(* IEC 61131-3 sources: rusty/tests/lit/single/polymorphism/interfaces/properties, 10 files *)

(* ---- basic_get_set.st ---- *)
// RUN: %COMPILE %s && %RUN | %CHECK %s
// Scenario: Single interface with a property declaring both PROPERTY_GET and PROPERTY_SET, implemented by a single
// function block. Assign the concrete instance to an interface variable and exercise both accessors
// through it. Baseline sanity test for property dispatch through interfaces.

INTERFACE IValue
    PROPERTY_GET value: DINT END_PROPERTY
    PROPERTY_SET value: DINT END_PROPERTY
END_INTERFACE

FUNCTION_BLOCK FbStore IMPLEMENTS IValue
    VAR
        _val : DINT := 10;
    END_VAR

    PROPERTY_GET value: DINT
        value := _val;
    END_PROPERTY

    PROPERTY_SET value: DINT
        _val := value;
    END_PROPERTY
END_FUNCTION_BLOCK

FUNCTION main
    VAR
        instance : FbStore;
        iface : IValue;
    END_VAR

    iface := instance;

    // CHECK: value=10
    printf('value=%d$N', iface.value);

    iface.value := 42;

    // CHECK-NEXT: value=42
    printf('value=%d$N', iface.value);

    iface.value := iface.value + 8;

    // CHECK-NEXT: value=50
    printf('value=%d$N', iface.value);
END_FUNCTION

(* ---- deep_chain_alternating_overrides.st ---- *)
// RUN: %COMPILE %s && %RUN | %CHECK %s
// Scenario: Three-level POU chain FbC → FbB → FbA, where FbA implements IValue. FbB overrides
// only the getter (adds 1000), FbC overrides only the setter (adds 2000). Dispatch through the
// interface should resolve each accessor to the most-derived override:
//   FbA → (FbA.get, FbA.set)
//   FbB → (FbB.get, FbA.set)
//   FbC → (FbB.get, FbC.set)

INTERFACE IValue
    PROPERTY_GET value: DINT END_PROPERTY
    PROPERTY_SET value: DINT END_PROPERTY
END_INTERFACE

FUNCTION_BLOCK FbA IMPLEMENTS IValue
    VAR
        _val : DINT := 10;
    END_VAR

    PROPERTY_GET value: DINT
        value := _val;
    END_PROPERTY

    PROPERTY_SET value: DINT
        _val := value;
    END_PROPERTY
END_FUNCTION_BLOCK

FUNCTION_BLOCK FbB EXTENDS FbA
    // Override only getter — adds 1000
    PROPERTY_GET value: DINT
        value := _val + 1000;
    END_PROPERTY
END_FUNCTION_BLOCK

FUNCTION_BLOCK FbC EXTENDS FbB
    // Override only setter — adds 2000
    PROPERTY_SET value: DINT
        _val := value + 2000;
    END_PROPERTY
END_FUNCTION_BLOCK

FUNCTION main
    VAR
        instanceA : FbA;
        instanceB : FbB;
        instanceC : FbC;
        iface : IValue;
    END_VAR

    // FbA: get=FbA, set=FbA
    iface := instanceA;
    printf('value=%d$N', iface.value);      // CHECK: value=10
    iface.value := 50;
    printf('value=%d$N', iface.value);      // CHECK-NEXT: value=50

    // FbB: get=FbB(+1000), set=FbA(inherited)
    iface := instanceB;
    printf('value=%d$N', iface.value);      // CHECK-NEXT: value=1010
    iface.value := 50;
    printf('value=%d$N', iface.value);      // CHECK-NEXT: value=1050

    // FbC: get=FbB(inherited, +1000), set=FbC(+2000)
    iface := instanceC;
    printf('value=%d$N', iface.value);      // CHECK-NEXT: value=1010
    iface.value := 50;
    printf('value=%d$N', iface.value);      // CHECK-NEXT: value=3050
END_FUNCTION

(* ---- diamond_hierarchy.st ---- *)
// RUN: %COMPILE %s && %RUN | %CHECK %s
// Scenario: Classic diamond pattern with a property at the root.
//     IA (property value)
//    /  \
//   IB   IC
//    \  /
//     ID
// IB adds method bar, IC adds method baz, ID adds method qux. A single function block
// FbImpl implements ID (and thus transitively IA, IB, IC). Dispatch through IA, IB, IC
// and ID variables should all resolve the property correctly, and each interface level
// should expose its respective methods.

INTERFACE IA
    PROPERTY_GET value: DINT END_PROPERTY
    PROPERTY_SET value: DINT END_PROPERTY
END_INTERFACE

INTERFACE IB EXTENDS IA
    METHOD bar END_METHOD
END_INTERFACE

INTERFACE IC EXTENDS IA
    METHOD baz END_METHOD
END_INTERFACE

INTERFACE ID EXTENDS IB, IC
    METHOD qux END_METHOD
END_INTERFACE

FUNCTION_BLOCK FbImpl IMPLEMENTS ID
    VAR
        _val : DINT := 10;
    END_VAR

    PROPERTY_GET value: DINT
        value := _val;
    END_PROPERTY

    PROPERTY_SET value: DINT
        _val := value;
    END_PROPERTY

    METHOD bar
        printf('bar(%d)$N', _val);
    END_METHOD

    METHOD baz
        printf('baz(%d)$N', _val);
    END_METHOD

    METHOD qux
        printf('qux(%d)$N', _val);
    END_METHOD
END_FUNCTION_BLOCK

FUNCTION main
    VAR
        instA : FbImpl;
        instB : FbImpl;
        instC : FbImpl;
        instD : FbImpl;
        refA : IA;
        refB : IB;
        refC : IC;
        refD : ID;
    END_VAR

    // Through IA — property only
    refA := instA;
    printf('value=%d$N', refA.value);           // CHECK: value=10
    refA.value := 42;
    printf('value=%d$N', refA.value);           // CHECK-NEXT: value=42

    // Through IB — property + bar
    refB := instB;
    printf('value=%d$N', refB.value);           // CHECK-NEXT: value=10
    refB.bar();                                 // CHECK-NEXT: bar(10)
    refB.value := 42;
    refB.bar();                                 // CHECK-NEXT: bar(42)
    printf('value=%d$N', refB.value);           // CHECK-NEXT: value=42

    // Through IC — property + baz
    refC := instC;
    printf('value=%d$N', refC.value);           // CHECK-NEXT: value=10
    refC.baz();                                 // CHECK-NEXT: baz(10)
    refC.value := 42;
    refC.baz();                                 // CHECK-NEXT: baz(42)
    printf('value=%d$N', refC.value);           // CHECK-NEXT: value=42

    // Through ID — property + bar + baz + qux
    refD := instD;
    printf('value=%d$N', refD.value);           // CHECK-NEXT: value=10
    refD.bar();                                 // CHECK-NEXT: bar(10)
    refD.baz();                                 // CHECK-NEXT: baz(10)
    refD.qux();                                 // CHECK-NEXT: qux(10)
    refD.value := 99;
    printf('value=%d$N', refD.value);           // CHECK-NEXT: value=99
    refD.bar();                                 // CHECK-NEXT: bar(99)
    refD.baz();                                 // CHECK-NEXT: baz(99)
    refD.qux();                                 // CHECK-NEXT: qux(99)
END_FUNCTION

(* ---- implicit_obligation_through_pou_chain.st ---- *)
// RUN: %COMPILE %s && %RUN | %CHECK %s
// Scenario: FbB extends FbA (which implements IValue) without overriding anything. FbC extends FbB,
// also without overriding. All three should be assignable to an IValue variable and dispatch
// correctly to FbA's inherited property accessors.

INTERFACE IValue
    PROPERTY_GET value: DINT END_PROPERTY
    PROPERTY_SET value: DINT END_PROPERTY
END_INTERFACE

FUNCTION_BLOCK FbA IMPLEMENTS IValue
    VAR
        _val : DINT := 10;
    END_VAR

    PROPERTY_GET value: DINT
        value := _val;
    END_PROPERTY

    PROPERTY_SET value: DINT
        _val := value;
    END_PROPERTY
END_FUNCTION_BLOCK

FUNCTION_BLOCK FbB EXTENDS FbA
    // No override — inherits everything from FbA
END_FUNCTION_BLOCK

FUNCTION_BLOCK FbC EXTENDS FbB
    // No override — inherits transitively from FbA
END_FUNCTION_BLOCK

FUNCTION main
    VAR
        instanceA : FbA;
        instanceB : FbB;
        instanceC : FbC;
        iface : IValue;
    END_VAR

    // FbA — direct implementor
    iface := instanceA;
    printf('value=%d$N', iface.value);      // CHECK: value=10
    iface.value := 42;
    printf('value=%d$N', iface.value);      // CHECK-NEXT: value=42

    // FbB — inherits from FbA (one level)
    iface := instanceB;
    printf('value=%d$N', iface.value);      // CHECK-NEXT: value=10
    iface.value := 77;
    printf('value=%d$N', iface.value);      // CHECK-NEXT: value=77

    // FbC — inherits transitively through FbB (two levels)
    iface := instanceC;
    printf('value=%d$N', iface.value);      // CHECK-NEXT: value=10
    iface.value := 99;
    printf('value=%d$N', iface.value);      // CHECK-NEXT: value=99
END_FUNCTION

(* ---- inherited_getter_overridden_setter.st ---- *)
// RUN: %COMPILE %s && %RUN | %CHECK %s
// Scenario: FbB extends FbA which implements interface IA with a PROPERTY_GET+PROPERTY_SET property. FbB overrides
// only the setter (adds 1000). Dispatch through an IA variable should use FbA's inherited getter
// and FbB's overridden setter when pointing at FbB.

INTERFACE IValue
    PROPERTY_GET value: DINT END_PROPERTY
    PROPERTY_SET value: DINT END_PROPERTY
END_INTERFACE

FUNCTION_BLOCK FbA IMPLEMENTS IValue
    VAR
        _val : DINT := 10;
    END_VAR

    PROPERTY_GET value: DINT
        value := _val;
    END_PROPERTY

    PROPERTY_SET value: DINT
        _val := value;
    END_PROPERTY
END_FUNCTION_BLOCK

FUNCTION_BLOCK FbB EXTENDS FbA
    // Override only setter — adds 1000 to distinguish
    PROPERTY_SET value: DINT
        _val := value + 1000;
    END_PROPERTY
END_FUNCTION_BLOCK

FUNCTION main
    VAR
        instanceA : FbA;
        instanceB : FbB;
        iface : IValue;
    END_VAR

    // FbA — both accessors from FbA
    iface := instanceA;
    printf('value=%d$N', iface.value);      // CHECK: value=10
    iface.value := 42;
    printf('value=%d$N', iface.value);      // CHECK-NEXT: value=42

    // FbB — getter inherited from FbA, setter overridden in FbB (+1000)
    iface := instanceB;
    printf('value=%d$N', iface.value);      // CHECK-NEXT: value=10
    iface.value := 42;
    printf('value=%d$N', iface.value);      // CHECK-NEXT: value=1042
END_FUNCTION

(* ---- inherited_setter_overridden_getter.st ---- *)
// RUN: %COMPILE %s && %RUN | %CHECK %s
// Scenario: FbB extends FbA which implements interface IA with a PROPERTY_GET+PROPERTY_SET property. FbB overrides
// only the getter (adds 1000). Dispatch through an IA variable should use FbB's overridden getter
// and FbA's inherited setter when pointing at FbB.

INTERFACE IValue
    PROPERTY_GET value: DINT END_PROPERTY
    PROPERTY_SET value: DINT END_PROPERTY
END_INTERFACE

FUNCTION_BLOCK FbA IMPLEMENTS IValue
    VAR
        _val : DINT := 10;
    END_VAR

    PROPERTY_GET value: DINT
        value := _val;
    END_PROPERTY

    PROPERTY_SET value: DINT
        _val := value;
    END_PROPERTY
END_FUNCTION_BLOCK

FUNCTION_BLOCK FbB EXTENDS FbA
    // Override only getter — adds 1000 to distinguish
    PROPERTY_GET value: DINT
        value := _val + 1000;
    END_PROPERTY
END_FUNCTION_BLOCK

FUNCTION main
    VAR
        instanceA : FbA;
        instanceB : FbB;
        iface : IValue;
    END_VAR

    // FbA — both accessors from FbA
    iface := instanceA;
    printf('value=%d$N', iface.value);      // CHECK: value=10
    iface.value := 42;
    printf('value=%d$N', iface.value);      // CHECK-NEXT: value=42

    // FbB — getter overridden in FbB (+1000), setter inherited from FbA
    iface := instanceB;
    printf('value=%d$N', iface.value);      // CHECK-NEXT: value=1010
    iface.value := 42;
    printf('value=%d$N', iface.value);      // CHECK-NEXT: value=1042
END_FUNCTION

(* ---- interface_hierarchy.st ---- *)
// RUN: %COMPILE %s && %RUN | %CHECK %s
// Scenario: IB extends IA, where IA declares a property and IB adds a method. FbImpl implements
// IB with both, FbChild extends FbImpl and overrides only the setter (adds 500). Dispatch through
// both IA and IB variables should resolve the property identically, while the method is only
// accessible through IB.

INTERFACE IA
    PROPERTY_GET value: DINT END_PROPERTY
    PROPERTY_SET value: DINT END_PROPERTY
END_INTERFACE

INTERFACE IB EXTENDS IA
    METHOD describe END_METHOD
END_INTERFACE

FUNCTION_BLOCK FbImpl IMPLEMENTS IB
    VAR
        _val : DINT := 10;
    END_VAR

    PROPERTY_GET value: DINT
        value := _val;
    END_PROPERTY

    PROPERTY_SET value: DINT
        _val := value;
    END_PROPERTY

    METHOD describe
        printf('FbImpl(%d)$N', _val);
    END_METHOD
END_FUNCTION_BLOCK

FUNCTION_BLOCK FbChild EXTENDS FbImpl
    // Override only setter — adds 500
    PROPERTY_SET value: DINT
        _val := value + 500;
    END_PROPERTY

    METHOD describe
        printf('FbChild(%d)$N', _val);
    END_METHOD
END_FUNCTION_BLOCK

FUNCTION main
    VAR
        implForA : FbImpl;
        implForB : FbImpl;
        childForA : FbChild;
        childForB : FbChild;
        refA : IA;
        refB : IB;
    END_VAR

    // Through IA — property only
    refA := implForA;
    printf('value=%d$N', refA.value);           // CHECK: value=10
    refA.value := 42;
    printf('value=%d$N', refA.value);           // CHECK-NEXT: value=42

    refA := childForA;
    printf('value=%d$N', refA.value);           // CHECK-NEXT: value=10
    refA.value := 42;
    printf('value=%d$N', refA.value);           // CHECK-NEXT: value=542

    // Through IB — property + method
    refB := implForB;
    refB.describe();                            // CHECK-NEXT: FbImpl(10)
    printf('value=%d$N', refB.value);           // CHECK-NEXT: value=10
    refB.value := 42;
    refB.describe();                            // CHECK-NEXT: FbImpl(42)

    refB := childForB;
    refB.describe();                            // CHECK-NEXT: FbChild(10)
    printf('value=%d$N', refB.value);           // CHECK-NEXT: value=10
    refB.value := 42;
    refB.describe();                            // CHECK-NEXT: FbChild(542)
    printf('value=%d$N', refB.value);           // CHECK-NEXT: value=542
END_FUNCTION

(* ---- mixed_methods_and_properties.st ---- *)
// RUN: %COMPILE %s && %RUN | %CHECK %s
// Scenario: An interface declares both a regular method and a property. Two function blocks
// implement the interface with different behaviors. Both the method and property are dispatched
// through the same interface variable, verifying they coexist cleanly in the itable.

INTERFACE IWidget
    METHOD describe END_METHOD

    PROPERTY_GET label: DINT END_PROPERTY
    PROPERTY_SET label: DINT END_PROPERTY
END_INTERFACE

FUNCTION_BLOCK FbButton IMPLEMENTS IWidget
    VAR
        _label : DINT := 1;
    END_VAR

    METHOD describe
        printf('Button(%d)$N', _label);
    END_METHOD

    PROPERTY_GET label: DINT
        label := _label;
    END_PROPERTY

    PROPERTY_SET label: DINT
        _label := label;
    END_PROPERTY
END_FUNCTION_BLOCK

FUNCTION_BLOCK FbSlider IMPLEMENTS IWidget
    VAR
        _label : DINT := 2;
    END_VAR

    METHOD describe
        printf('Slider(%d)$N', _label);
    END_METHOD

    PROPERTY_GET label: DINT
        label := _label * 10;
    END_PROPERTY

    PROPERTY_SET label: DINT
        _label := label + 100;
    END_PROPERTY
END_FUNCTION_BLOCK

FUNCTION main
    VAR
        button : FbButton;
        slider : FbSlider;
        iface : IWidget;
    END_VAR

    // FbButton
    iface := button;
    iface.describe();                           // CHECK: Button(1)
    printf('label=%d$N', iface.label);          // CHECK-NEXT: label=1
    iface.label := 42;
    iface.describe();                           // CHECK-NEXT: Button(42)
    printf('label=%d$N', iface.label);          // CHECK-NEXT: label=42

    // FbSlider — getter returns _label * 10, setter stores label + 100
    iface := slider;
    iface.describe();                           // CHECK-NEXT: Slider(2)
    printf('label=%d$N', iface.label);          // CHECK-NEXT: label=20
    iface.label := 99;
    iface.describe();                           // CHECK-NEXT: Slider(199)
    printf('label=%d$N', iface.label);          // CHECK-NEXT: label=1990
END_FUNCTION

(* ---- multiple_implementors.st ---- *)
// RUN: %COMPILE %s && %RUN | %CHECK %s
// Scenario: Two function blocks implement the same interface property with different backing logic.
// FbPlain returns the stored value directly, FbDoubling returns twice the stored value. Assigning
// each to the same interface variable and reading the property verifies that dispatch picks the
// correct accessor implementation each time.

INTERFACE IValue
    PROPERTY_GET value: DINT END_PROPERTY
    PROPERTY_SET value: DINT END_PROPERTY
END_INTERFACE

FUNCTION_BLOCK FbPlain IMPLEMENTS IValue
    VAR
        _val : DINT := 10;
    END_VAR

    PROPERTY_GET value: DINT
        value := _val;
    END_PROPERTY

    PROPERTY_SET value: DINT
        _val := value;
    END_PROPERTY
END_FUNCTION_BLOCK

FUNCTION_BLOCK FbDoubling IMPLEMENTS IValue
    VAR
        _val : DINT := 10;
    END_VAR

    PROPERTY_GET value: DINT
        value := _val * 2;
    END_PROPERTY

    PROPERTY_SET value: DINT
        _val := value;
    END_PROPERTY
END_FUNCTION_BLOCK

FUNCTION main
    VAR
        plain : FbPlain;
        doubling : FbDoubling;
        iface : IValue;
    END_VAR

    // FbPlain — getter returns _val directly
    iface := plain;
    printf('value=%d$N', iface.value);      // CHECK: value=10
    iface.value := 42;
    printf('value=%d$N', iface.value);      // CHECK-NEXT: value=42

    // FbDoubling — getter returns _val * 2
    iface := doubling;
    printf('value=%d$N', iface.value);      // CHECK-NEXT: value=20
    iface.value := 42;
    printf('value=%d$N', iface.value);      // CHECK-NEXT: value=84
END_FUNCTION

(* ---- property_get_as_function_argument.st ---- *)
// RUN: %COMPILE %s && %RUN | %CHECK %s
// Scenario: Passing a property getter result as an argument to a function, dispatched through
// an interface reference. Mirrors the `property_get_as_function_argument` unit test.

INTERFACE IValue
    PROPERTY_GET value: DINT END_PROPERTY
END_INTERFACE

FUNCTION_BLOCK FbStore IMPLEMENTS IValue
    VAR
        _val : DINT;
    END_VAR

    PROPERTY_GET value: DINT
        value := _val;
    END_PROPERTY
END_FUNCTION_BLOCK

FUNCTION consumer
    VAR_INPUT
        x : DINT;
    END_VAR

    printf('consumed=%d$N', x);
END_FUNCTION

FUNCTION main
    VAR
        instance : FbStore;
        iface : IValue;
    END_VAR

    instance._val := 42;
    iface := instance;

    // Property getter result passed directly as function argument
    consumer(iface.value);              // CHECK: consumed=42

    instance._val := 99;
    iface := instance;
    consumer(iface.value);              // CHECK-NEXT: consumed=99
END_FUNCTION
